(* IEC 61131-3 sources: sigmatek-logger-api/IXON_API/Network/IXON_Log, 1 file *)

(* ---- ONE_IXON_Log_Table.st ---- *)
#define OBJECTS_CONFIG

//Define part of class _TCPIPClient
#define TCPCLT_ERROR_NO            0
  #define TCPCLT_ERROR_INVALID_SOCK  -1
  #define TCPCLT_ERROR_CONNECTION    -2
  #define TCPCLT_ERROR_TIMEOUT       -3

  #define TCP_CLT_SEND_OK               0
  #define TCP_CLT_INVALID_HANDLE        -1
  #define TCP_CLT_NOT_CONNECTED         -2
  #define TCP_CLT_SEND_FAILED           -3
  #define TCP_CLT_SEND_BUFFER_FULL      -4
  #define TCP_CLT_DATA_TO_BIG_FOR_DIRECT_SENDING   -5
  #define TCP_CLT_MAXLEN_SEMANAME     32

  #define TCP_CLT_ERR_SET_PARA_INVALID_CMD     -10
  #define TCP_CLT_ERR_SET_PARA_INVALID_SUB_CMD -11

  #define TCP_CLT_ERR_TASK_ALREADY_EXIST       -12

  #define TCP_CLT_ERR_SET_PARA_CMD_NOT_SUPPORTED  -13

  #ifndef OS_VERSION_MIN_SALAMANDER
    #define OS_VERSION_MIN_SALAMANDER          0x9000
  #endif

  #define TCP_CLT_NO_ERROR                          0

  // - RETURN VALUES PRIVATE METHOD Read_LSLOBJ_CRC32
  #define TCP_CLT_ERR_GET_LSLOBJ_NAME             -20
  #define TCP_CLT_ERR_INVALID_POINTER             -21

  // - RETURN VALUES PRIVATE METHOD Read_AP_TaskPeriod
  #define TCP_CLT_ERR_TASK_TIME_NO_APP            -31
  #define TCP_CLT_ERR_TASK_TIME_WRONG_TASK_TYPE   -33
  #define TCP_CLT_ERR_TASK_TIME_OBJ_NOT_FOUND     -35

  // - RETURN VALUES PRIVATE METHOD AP_TaskCreate
  #define TCP_CLT_ERR_TASK_CREATE                 -40

  // - RETURN VALUES PRIVATE METHOD AP_SemaCreate
  #define TCP_CLT_ERR_SEMA_CREATE                 -50
  #define TCP_CLT_ERR_SEMA_INVALID_IDX            -51
  #define TCP_CLT_ERR_SEMA_INVALID_NAME           -52

  #define TCP_CLT_SEND_BUFFER_EMPTY                -6
  #define TCP_CLT_ERR_SEND_BUFFER_FATAL_ERROR      -7

  #define TCP_CLT_ERR_NO_SSL_INTERFACE             -8
  #define TCP_CLT_ERR_NO_TCP_INTERFACE             -9

  #define TCP_CLT_ERR_INVALID_PARA_TCP            -60
  #define TCP_CLT_ERR_INVALID_PARA_SSL            -61

  #define TCP_CLT_ERR_CONN_MEMORY                 -70
  #define TCP_CLT_ERR_MAX_CONN                    -80
  #define TCP_CLT_ERR_MAIN_INIT                   -90

  #define TCP_CLT_ERR_GROUP_OS                      0
  #define TCP_CLT_ERR_GROUP_AP                      1

  #define TCP_CLT_ERR_CODE_AP_TIMEOUT              -1

  #ifndef INIT_FIRSTSCAN
    #define INIT_FIRSTSCAN                         12
  #endif

  #ifndef AP_TASK_PRIORITY_DEFAULT
    #define AP_TASK_PRIORITY_DEFAULT               14
  #endif

  #define TCP_CLT_CMD_KEEP_ALIVE_PARA               2
  #define TCP_CLT_SUB_CMD_KEEP_ALIVE_INTERVAL       0
  #define TCP_CLT_SUB_CMD_KEEP_ALIVE_RETRY          1
  #define TCP_CLT_SUB_CMD_KEEP_ALIVE_TIMEOUT        2

  #define TCP_CLT_INFO_DISCONNECT                   0
  #define TCP_CLT_INFO_CONNECT                      1
  #define TCP_CLT_INFO_DELETED                      2

  #ifndef KEEPALIVE_INTERVAL_DEFAULT
    #define KEEPALIVE_INTERVAL_DEFAULT           7200
  #endif

  #ifndef KEEPALIVE_RETRYTIME_DEFAULT
    #define KEEPALIVE_RETRYTIME_DEFAULT            75
  #endif

  #ifndef KEEPALIVE_RETRYCNT_DEFUALT
    #define KEEPALIVE_RETRYCNT_DEFUALT             10
  #endif

  #ifndef CLOSE_SOCKET_TYPE_DEFAULT
    #define CLOSE_SOCKET_TYPE_DEFAULT               0
  #endif
#include "..\..\Class\_TCPIPClient\_TCPIPClient.h"
#include "..\..\Class\_TCPIPClient\SalamanderDelay.h"
#include "..\..\Class\_TCPIPClient\lsl_st_ssl_user.h"
//Define part of class cIXONConv10Value
#DEFINE MAX_NAME_LENGTH 100
#DEFINE MAX_VALUE_LENGTH 10
#DEFINE MAX_DATASTRING_LENGTH 1024
//Define part of class cIXONConv5Int5Str
#DEFINE MAX_NAME_LENGTH 100
#DEFINE MAX_INTEGER_LENGTH 10
#DEFINE MAX_DATASTRING_LENGTH 1024
#DEFINE MAX_STRING_LENGTH 100
//Define part of class IXON_LoggerAPI_Interface
#define SND_DATA_ARRAY_SIZE 1024
#define SND_ARRAY_SIZE 20
#define RCV_DATA_ARRAY_SIZE 1024
#include <.\lsl_st_mt.h>

FUNCTION GLOBAL TAB ONE_IXON_Log
-1$UINT, 0$UINT,
0$UINT, 0$UINT,

12$UDINT,
TO_UDINT(916194998), "_CheckSum", 1$UINT, 0$UINT, 1$UINT,
TO_UDINT(1778057824), "_TCPIPClient", 1$UINT, 1$UINT, 1$UINT,
TO_UDINT(670188634), "_TCPIPClientInterface", 1$UINT, 1$UINT, 0$UINT,
TO_UDINT(2199147857), "cIXONConv10Value", 0$UINT, 0$UINT, 1$UINT,
TO_UDINT(2966690256), "cIXONConv5Int5Str", 0$UINT, 0$UINT, 1$UINT,
TO_UDINT(2366984241), "IXON_LoggerAPI", 0$UINT, 0$UINT, 1$UINT,
TO_UDINT(357781282), "IXON_LoggerAPI_Interface", 0$UINT, 0$UINT, 1$UINT,
TO_UDINT(2225119864), "MerkerEx", 1$UINT, 22$UINT, 33$UINT,
TO_UDINT(3963750506), "Pulse", 0$UINT, 0$UINT, 1$UINT,
TO_UDINT(1850111279), "String", 1$UINT, 11$UINT, 33$UINT,
TO_UDINT(2898603620), "StringInternal", 1$UINT, 84$UINT, 0$UINT,
TO_UDINT(3232495061), "VirtualBaseInit", 1$UINT, 3$UINT, 0$UINT,

1$UINT, TO_UDINT(3180115317), "IXON_LOGGERAPI1\_TCPIPCLIENT1\CHECKSUM",

1$UINT, TO_UDINT(1796594274), "IXON_LOGGERAPI1\_TCPIPCLIENT1",

_NO_ATTR, TO_UDINT(3085999121), "GRIPPERSIXONLOG",

_NO_ATTR, TO_UDINT(1798062204), "BATCHIXONLOG",

_NO_ATTR, TO_UDINT(3532651229), "IXON_LOGGERAPI1",

1$UINT, TO_UDINT(1003265729), "IXON_LOGGERAPI1\MYTCPIPCLIENT1",

1$UINT, TO_UDINT(3192771373), "BATCHIXONLOG\INTEGERNAME1\MERKEREX0",
1$UINT, TO_UDINT(665826604), "BATCHIXONLOG\INTEGERNAME2\MERKEREX0",
1$UINT, TO_UDINT(3860949740), "BATCHIXONLOG\INTEGERNAME3\MERKEREX0",
1$UINT, TO_UDINT(3474620271), "BATCHIXONLOG\INTEGERNAME4\MERKEREX0",
1$UINT, TO_UDINT(244621487), "BATCHIXONLOG\INTEGERNAME5\MERKEREX0",
1$UINT, TO_UDINT(2181923968), "BATCHIXONLOG\STRING1\MERKEREX0",
1$UINT, TO_UDINT(468705921), "BATCHIXONLOG\STRING2\MERKEREX0",
1$UINT, TO_UDINT(3663805761), "BATCHIXONLOG\STRING3\MERKEREX0",
1$UINT, TO_UDINT(4082772162), "BATCHIXONLOG\STRING4\MERKEREX0",
1$UINT, TO_UDINT(852817666), "BATCHIXONLOG\STRING5\MERKEREX0",
1$UINT, TO_UDINT(2342531462), "BATCHIXONLOG\STRINGNAME1\MERKEREX0",
1$UINT, TO_UDINT(306337671), "BATCHIXONLOG\STRINGNAME2\MERKEREX0",
1$UINT, TO_UDINT(3553396807), "BATCHIXONLOG\STRINGNAME3\MERKEREX0",
1$UINT, TO_UDINT(4210531780), "BATCHIXONLOG\STRINGNAME4\MERKEREX0",
1$UINT, TO_UDINT(997802500), "BATCHIXONLOG\STRINGNAME5\MERKEREX0",
1$UINT, TO_UDINT(2779010355), "BATCHIXONLOG\TRIGGERNAME\MERKEREX0",
1$UINT, TO_UDINT(4245150780), "GRIPPERSIXONLOG\NAME10\MERKEREX0",
1$UINT, TO_UDINT(2566426530), "GRIPPERSIXONLOG\NAME1\MERKEREX0",
1$UINT, TO_UDINT(18540963), "GRIPPERSIXONLOG\NAME2\MERKEREX0",
1$UINT, TO_UDINT(3230938723), "GRIPPERSIXONLOG\NAME3\MERKEREX0",
1$UINT, TO_UDINT(3920569312), "GRIPPERSIXONLOG\NAME4\MERKEREX0",
1$UINT, TO_UDINT(673315872), "GRIPPERSIXONLOG\NAME5\MERKEREX0",
1$UINT, TO_UDINT(2982386209), "GRIPPERSIXONLOG\NAME6\MERKEREX0",
1$UINT, TO_UDINT(1884112353), "GRIPPERSIXONLOG\NAME7\MERKEREX0",
1$UINT, TO_UDINT(3820335399), "GRIPPERSIXONLOG\NAME8\MERKEREX0",
1$UINT, TO_UDINT(574320359), "GRIPPERSIXONLOG\NAME9\MERKEREX0",
1$UINT, TO_UDINT(3865678693), "GRIPPERSIXONLOG\TRIGGERNAME\MERKEREX0",
1$UINT, TO_UDINT(2981893656), "IXON_LOGGERAPI1\MYTCPIPCLIENT1\ST_IPADDRIXON\MERKEREX0",
1$UINT, TO_UDINT(2486479070), "IXON_LOGGERAPI1\MYTCPIPCLIENT1\ST_IPADDRPLC\MERKEREX0",
1$UINT, TO_UDINT(3086082301), "IXON_LOGGERAPI1\MYTCPIPCLIENT1\ST_PASSWORDIXON\MERKEREX0",
1$UINT, TO_UDINT(3369279868), "IXON_LOGGERAPI1\_TCPIPCLIENT1\STRSEMANAME01\MERKEREX0",
1$UINT, TO_UDINT(1362184061), "IXON_LOGGERAPI1\_TCPIPCLIENT1\STRSEMANAME02\MERKEREX0",
1$UINT, TO_UDINT(3451953391), "IXON_LOGGERAPI1\_TCPIPCLIENT1\STRTASKNAME\MERKEREX0",

_NO_ATTR, TO_UDINT(777463289), "PULSE1",

1$UINT, TO_UDINT(808633261), "BATCHIXONLOG\INTEGERNAME1",
1$UINT, TO_UDINT(2839253527), "BATCHIXONLOG\INTEGERNAME2",
1$UINT, TO_UDINT(3728515713), "BATCHIXONLOG\INTEGERNAME3",
1$UINT, TO_UDINT(1079523106), "BATCHIXONLOG\INTEGERNAME4",
1$UINT, TO_UDINT(928974772), "BATCHIXONLOG\INTEGERNAME5",
1$UINT, TO_UDINT(4091281586), "BATCHIXONLOG\STRING1",
1$UINT, TO_UDINT(1792364808), "BATCHIXONLOG\STRING2",
1$UINT, TO_UDINT(500326814), "BATCHIXONLOG\STRING3",
1$UINT, TO_UDINT(2209805373), "BATCHIXONLOG\STRING4",
1$UINT, TO_UDINT(4105290923), "BATCHIXONLOG\STRING5",
1$UINT, TO_UDINT(1673436439), "BATCHIXONLOG\STRINGNAME1",
1$UINT, TO_UDINT(4206349485), "BATCHIXONLOG\STRINGNAME2",
1$UINT, TO_UDINT(2377186363), "BATCHIXONLOG\STRINGNAME3",
1$UINT, TO_UDINT(332687768), "BATCHIXONLOG\STRINGNAME4",
1$UINT, TO_UDINT(1691572494), "BATCHIXONLOG\STRINGNAME5",
1$UINT, TO_UDINT(3473702409), "BATCHIXONLOG\TRIGGERNAME",
1$UINT, TO_UDINT(813494443), "GRIPPERSIXONLOG\NAME1",
1$UINT, TO_UDINT(3052394929), "GRIPPERSIXONLOG\NAME10",
1$UINT, TO_UDINT(2843058449), "GRIPPERSIXONLOG\NAME2",
1$UINT, TO_UDINT(3732050311), "GRIPPERSIXONLOG\NAME3",
1$UINT, TO_UDINT(1075184676), "GRIPPERSIXONLOG\NAME4",
1$UINT, TO_UDINT(923874482), "GRIPPERSIXONLOG\NAME5",
1$UINT, TO_UDINT(2920834312), "GRIPPERSIXONLOG\NAME6",
1$UINT, TO_UDINT(3642709406), "GRIPPERSIXONLOG\NAME7",
1$UINT, TO_UDINT(1235240975), "GRIPPERSIXONLOG\NAME8",
1$UINT, TO_UDINT(1051162777), "GRIPPERSIXONLOG\NAME9",
1$UINT, TO_UDINT(3416962169), "GRIPPERSIXONLOG\TRIGGERNAME",
1$UINT, TO_UDINT(2721538750), "IXON_LOGGERAPI1\MYTCPIPCLIENT1\ST_IPADDRIXON",
1$UINT, TO_UDINT(1805041610), "IXON_LOGGERAPI1\MYTCPIPCLIENT1\ST_IPADDRPLC",
1$UINT, TO_UDINT(1852407263), "IXON_LOGGERAPI1\MYTCPIPCLIENT1\ST_PASSWORDIXON",
1$UINT, TO_UDINT(962394143), "IXON_LOGGERAPI1\_TCPIPCLIENT1\STRSEMANAME01",
1$UINT, TO_UDINT(2689968549), "IXON_LOGGERAPI1\_TCPIPCLIENT1\STRSEMANAME02",
1$UINT, TO_UDINT(2790321702), "IXON_LOGGERAPI1\_TCPIPCLIENT1\STRTASKNAME",

//Internal connections
0$UDINT,
69$UDINT,
TO_UDINT(1), "CheckSum", TO_UDINT(0),
TO_UDINT(1), "StrTaskName", TO_UDINT(72),
TO_UDINT(1), "StrSemaName01", TO_UDINT(70),
TO_UDINT(1), "StrSemaName02", TO_UDINT(71),
TO_UDINT(2), "Name3", TO_UDINT(59),
TO_UDINT(2), "Name2", TO_UDINT(58),
TO_UDINT(2), "Name1", TO_UDINT(56),
TO_UDINT(2), "Name4", TO_UDINT(60),
TO_UDINT(2), "Name5", TO_UDINT(61),
TO_UDINT(2), "Name6", TO_UDINT(62),
TO_UDINT(2), "Name7", TO_UDINT(63),
TO_UDINT(2), "Name8", TO_UDINT(64),
TO_UDINT(2), "Name9", TO_UDINT(65),
TO_UDINT(2), "Name10", TO_UDINT(57),
TO_UDINT(2), "TriggerName", TO_UDINT(66),
TO_UDINT(3), "TriggerName", TO_UDINT(55),
TO_UDINT(3), "String1", TO_UDINT(45),
TO_UDINT(3), "String2", TO_UDINT(46),
TO_UDINT(3), "String3", TO_UDINT(47),
TO_UDINT(3), "String4", TO_UDINT(48),
TO_UDINT(3), "String5", TO_UDINT(49),
TO_UDINT(3), "IntegerName1", TO_UDINT(40),
TO_UDINT(3), "IntegerName2", TO_UDINT(41),
TO_UDINT(3), "IntegerName3", TO_UDINT(42),
TO_UDINT(3), "IntegerName4", TO_UDINT(43),
TO_UDINT(3), "IntegerName5", TO_UDINT(44),
TO_UDINT(3), "StringName1", TO_UDINT(50),
TO_UDINT(3), "StringName2", TO_UDINT(51),
TO_UDINT(3), "StringName3", TO_UDINT(52),
TO_UDINT(3), "StringName4", TO_UDINT(53),
TO_UDINT(3), "StringName5", TO_UDINT(54),
TO_UDINT(4), "_TCPIPClient1", TO_UDINT(1),
TO_UDINT(4), "MyTCPIPClient1", TO_UDINT(5),
TO_UDINT(5), "ST_IPAddrIXON", TO_UDINT(67),
TO_UDINT(5), "ST_PasswordIXON", TO_UDINT(69),
TO_UDINT(5), "ST_IPAddrPLC", TO_UDINT(68),
TO_UDINT(40), "MerkerEx0", TO_UDINT(6),
TO_UDINT(41), "MerkerEx0", TO_UDINT(7),
TO_UDINT(42), "MerkerEx0", TO_UDINT(8),
TO_UDINT(43), "MerkerEx0", TO_UDINT(9),
TO_UDINT(44), "MerkerEx0", TO_UDINT(10),
TO_UDINT(45), "MerkerEx0", TO_UDINT(11),
TO_UDINT(46), "MerkerEx0", TO_UDINT(12),
TO_UDINT(47), "MerkerEx0", TO_UDINT(13),
TO_UDINT(48), "MerkerEx0", TO_UDINT(14),
TO_UDINT(49), "MerkerEx0", TO_UDINT(15),
TO_UDINT(50), "MerkerEx0", TO_UDINT(16),
TO_UDINT(51), "MerkerEx0", TO_UDINT(17),
TO_UDINT(52), "MerkerEx0", TO_UDINT(18),
TO_UDINT(53), "MerkerEx0", TO_UDINT(19),
TO_UDINT(54), "MerkerEx0", TO_UDINT(20),
TO_UDINT(55), "MerkerEx0", TO_UDINT(21),
TO_UDINT(56), "MerkerEx0", TO_UDINT(23),
TO_UDINT(57), "MerkerEx0", TO_UDINT(22),
TO_UDINT(58), "MerkerEx0", TO_UDINT(24),
TO_UDINT(59), "MerkerEx0", TO_UDINT(25),
TO_UDINT(60), "MerkerEx0", TO_UDINT(26),
TO_UDINT(61), "MerkerEx0", TO_UDINT(27),
TO_UDINT(62), "MerkerEx0", TO_UDINT(28),
TO_UDINT(63), "MerkerEx0", TO_UDINT(29),
TO_UDINT(64), "MerkerEx0", TO_UDINT(30),
TO_UDINT(65), "MerkerEx0", TO_UDINT(31),
TO_UDINT(66), "MerkerEx0", TO_UDINT(32),
TO_UDINT(67), "MerkerEx0", TO_UDINT(33),
TO_UDINT(68), "MerkerEx0", TO_UDINT(34),
TO_UDINT(69), "MerkerEx0", TO_UDINT(35),
TO_UDINT(70), "MerkerEx0", TO_UDINT(36),
TO_UDINT(71), "MerkerEx0", TO_UDINT(37),
TO_UDINT(72), "MerkerEx0", TO_UDINT(38),
0$UDINT,
39$UDINT,
TO_UDINT(2), "ToIXON_LoggerAPI", TO_UDINT(5), "ClassSvr",
TO_UDINT(3), "ToIXON_LoggerAPI", TO_UDINT(5), "ClassSvr",
TO_UDINT(5), "_TCPIPClient", TO_UDINT(1), "Control",
TO_UDINT(39), "PulseOut1", TO_UDINT(2), "sCmdConvert",
TO_UDINT(39), "PulseOut2", TO_UDINT(2), "sValue1",
TO_UDINT(39), "PulseOut3", TO_UDINT(3), "sCmdConvert",
TO_UDINT(40), "DataBuffer", TO_UDINT(6), "m_udLength",
TO_UDINT(41), "DataBuffer", TO_UDINT(7), "m_udLength",
TO_UDINT(42), "DataBuffer", TO_UDINT(8), "m_udLength",
TO_UDINT(43), "DataBuffer", TO_UDINT(9), "m_udLength",
TO_UDINT(44), "DataBuffer", TO_UDINT(10), "m_udLength",
TO_UDINT(45), "DataBuffer", TO_UDINT(11), "m_udLength",
TO_UDINT(46), "DataBuffer", TO_UDINT(12), "m_udLength",
TO_UDINT(47), "DataBuffer", TO_UDINT(13), "m_udLength",
TO_UDINT(48), "DataBuffer", TO_UDINT(14), "m_udLength",
TO_UDINT(49), "DataBuffer", TO_UDINT(15), "m_udLength",
TO_UDINT(50), "DataBuffer", TO_UDINT(16), "m_udLength",
TO_UDINT(51), "DataBuffer", TO_UDINT(17), "m_udLength",
TO_UDINT(52), "DataBuffer", TO_UDINT(18), "m_udLength",
TO_UDINT(53), "DataBuffer", TO_UDINT(19), "m_udLength",
TO_UDINT(54), "DataBuffer", TO_UDINT(20), "m_udLength",
TO_UDINT(55), "DataBuffer", TO_UDINT(21), "m_udLength",
TO_UDINT(56), "DataBuffer", TO_UDINT(23), "m_udLength",
TO_UDINT(57), "DataBuffer", TO_UDINT(22), "m_udLength",
TO_UDINT(58), "DataBuffer", TO_UDINT(24), "m_udLength",
TO_UDINT(59), "DataBuffer", TO_UDINT(25), "m_udLength",
TO_UDINT(60), "DataBuffer", TO_UDINT(26), "m_udLength",
TO_UDINT(61), "DataBuffer", TO_UDINT(27), "m_udLength",
TO_UDINT(62), "DataBuffer", TO_UDINT(28), "m_udLength",
TO_UDINT(63), "DataBuffer", TO_UDINT(29), "m_udLength",
TO_UDINT(64), "DataBuffer", TO_UDINT(30), "m_udLength",
TO_UDINT(65), "DataBuffer", TO_UDINT(31), "m_udLength",
TO_UDINT(66), "DataBuffer", TO_UDINT(32), "m_udLength",
TO_UDINT(67), "DataBuffer", TO_UDINT(33), "m_udLength",
TO_UDINT(68), "DataBuffer", TO_UDINT(34), "m_udLength",
TO_UDINT(69), "DataBuffer", TO_UDINT(35), "m_udLength",
TO_UDINT(70), "DataBuffer", TO_UDINT(36), "m_udLength",
TO_UDINT(71), "DataBuffer", TO_UDINT(37), "m_udLength",
TO_UDINT(72), "DataBuffer", TO_UDINT(38), "m_udLength",

//Initialization values
0$UDINT,
71$UDINT,
TO_UDINT(1), "Port", TO_UDINT(9230),//|IXON_Log.IXON_LoggerAPI1\_TCPIPClient1.Port;
TO_UDINT(1), "MaxConnections", TO_UDINT(0),//|IXON_Log.IXON_LoggerAPI1\_TCPIPClient1.MaxConnections;
TO_UDINT(2), "sSetInitNrOfEntrys", TO_UDINT(8),//|IXON_Log.GrippersIXONLog.sSetInitNrOfEntrys;
TO_UDINT(3), "sSetInitNrOfInteger", TO_UDINT(1),//|IXON_Log.BatchIXONLog.sSetInitNrOfInteger;
TO_UDINT(3), "sSetInitNrOfString", TO_UDINT(3),//|IXON_Log.BatchIXONLog.sSetInitNrOfString;
TO_UDINT(6), "ThreadSafe", TO_UDINT(0),//|IXON_Log.IntegerName1\BatchIXONLog\MerkerEx0.ThreadSafe;
TO_UDINT(7), "ThreadSafe", TO_UDINT(0),//|IXON_Log.IntegerName2\BatchIXONLog\MerkerEx0.ThreadSafe;
TO_UDINT(8), "ThreadSafe", TO_UDINT(0),//|IXON_Log.IntegerName3\BatchIXONLog\MerkerEx0.ThreadSafe;
TO_UDINT(9), "ThreadSafe", TO_UDINT(0),//|IXON_Log.IntegerName4\BatchIXONLog\MerkerEx0.ThreadSafe;
TO_UDINT(10), "ThreadSafe", TO_UDINT(0),//|IXON_Log.IntegerName5\BatchIXONLog\MerkerEx0.ThreadSafe;
TO_UDINT(11), "ThreadSafe", TO_UDINT(0),//|IXON_Log.String1\BatchIXONLog\MerkerEx0.ThreadSafe;
TO_UDINT(12), "ThreadSafe", TO_UDINT(0),//|IXON_Log.String2\BatchIXONLog\MerkerEx0.ThreadSafe;
TO_UDINT(13), "ThreadSafe", TO_UDINT(0),//|IXON_Log.String3\BatchIXONLog\MerkerEx0.ThreadSafe;
TO_UDINT(14), "ThreadSafe", TO_UDINT(0),//|IXON_Log.String4\BatchIXONLog\MerkerEx0.ThreadSafe;
TO_UDINT(15), "ThreadSafe", TO_UDINT(0),//|IXON_Log.String5\BatchIXONLog\MerkerEx0.ThreadSafe;
TO_UDINT(16), "ThreadSafe", TO_UDINT(0),//|IXON_Log.StringName1\BatchIXONLog\MerkerEx0.ThreadSafe;
TO_UDINT(17), "ThreadSafe", TO_UDINT(0),//|IXON_Log.StringName2\BatchIXONLog\MerkerEx0.ThreadSafe;
TO_UDINT(18), "ThreadSafe", TO_UDINT(0),//|IXON_Log.StringName3\BatchIXONLog\MerkerEx0.ThreadSafe;
TO_UDINT(19), "ThreadSafe", TO_UDINT(0),//|IXON_Log.StringName4\BatchIXONLog\MerkerEx0.ThreadSafe;
TO_UDINT(20), "ThreadSafe", TO_UDINT(0),//|IXON_Log.StringName5\BatchIXONLog\MerkerEx0.ThreadSafe;
TO_UDINT(21), "ThreadSafe", TO_UDINT(0),//|IXON_Log.TriggerName\BatchIXONLog\MerkerEx0.ThreadSafe;
TO_UDINT(22), "ThreadSafe", TO_UDINT(0),//|IXON_Log.Name10\GrippersIXONLog\MerkerEx0.ThreadSafe;
TO_UDINT(23), "ThreadSafe", TO_UDINT(0),//|IXON_Log.Name1\GrippersIXONLog\MerkerEx0.ThreadSafe;
TO_UDINT(24), "ThreadSafe", TO_UDINT(0),//|IXON_Log.Name2\GrippersIXONLog\MerkerEx0.ThreadSafe;
TO_UDINT(25), "ThreadSafe", TO_UDINT(0),//|IXON_Log.Name3\GrippersIXONLog\MerkerEx0.ThreadSafe;
TO_UDINT(26), "ThreadSafe", TO_UDINT(0),//|IXON_Log.Name4\GrippersIXONLog\MerkerEx0.ThreadSafe;
TO_UDINT(27), "ThreadSafe", TO_UDINT(0),//|IXON_Log.Name5\GrippersIXONLog\MerkerEx0.ThreadSafe;
TO_UDINT(28), "ThreadSafe", TO_UDINT(0),//|IXON_Log.Name6\GrippersIXONLog\MerkerEx0.ThreadSafe;
TO_UDINT(29), "ThreadSafe", TO_UDINT(0),//|IXON_Log.Name7\GrippersIXONLog\MerkerEx0.ThreadSafe;
TO_UDINT(30), "ThreadSafe", TO_UDINT(0),//|IXON_Log.Name8\GrippersIXONLog\MerkerEx0.ThreadSafe;
TO_UDINT(31), "ThreadSafe", TO_UDINT(0),//|IXON_Log.Name9\GrippersIXONLog\MerkerEx0.ThreadSafe;
TO_UDINT(32), "ThreadSafe", TO_UDINT(0),//|IXON_Log.TriggerName\GrippersIXONLog\MerkerEx0.ThreadSafe;
TO_UDINT(33), "ThreadSafe", TO_UDINT(0),//|IXON_Log.ST_IPAddrIXON\MyTCPIPClient1\IXON_LoggerAPI1\MerkerEx0.ThreadSafe;
TO_UDINT(34), "ThreadSafe", TO_UDINT(0),//|IXON_Log.ST_IPAddrPLC\MyTCPIPClient1\IXON_LoggerAPI1\MerkerEx0.ThreadSafe;
TO_UDINT(35), "ThreadSafe", TO_UDINT(0),//|IXON_Log.ST_PasswordIXON\MyTCPIPClient1\IXON_LoggerAPI1\MerkerEx0.ThreadSafe;
TO_UDINT(36), "ThreadSafe", TO_UDINT(0),//|IXON_Log.StrSemaName01\_TCPIPClient1\IXON_LoggerAPI1\MerkerEx0.ThreadSafe;
TO_UDINT(37), "ThreadSafe", TO_UDINT(0),//|IXON_Log.StrSemaName02\_TCPIPClient1\IXON_LoggerAPI1\MerkerEx0.ThreadSafe;
TO_UDINT(38), "ThreadSafe", TO_UDINT(0),//|IXON_Log.StrTaskName\_TCPIPClient1\IXON_LoggerAPI1\MerkerEx0.ThreadSafe;
TO_UDINT(40), "SingleRealloc", TO_UDINT(1),//|IXON_Log.BatchIXONLog\IntegerName1.SingleRealloc;
TO_UDINT(41), "SingleRealloc", TO_UDINT(1),//|IXON_Log.BatchIXONLog\IntegerName2.SingleRealloc;
TO_UDINT(42), "SingleRealloc", TO_UDINT(1),//|IXON_Log.BatchIXONLog\IntegerName3.SingleRealloc;
TO_UDINT(43), "SingleRealloc", TO_UDINT(1),//|IXON_Log.BatchIXONLog\IntegerName4.SingleRealloc;
TO_UDINT(44), "SingleRealloc", TO_UDINT(1),//|IXON_Log.BatchIXONLog\IntegerName5.SingleRealloc;
TO_UDINT(45), "SingleRealloc", TO_UDINT(1),//|IXON_Log.BatchIXONLog\String1.SingleRealloc;
TO_UDINT(46), "SingleRealloc", TO_UDINT(1),//|IXON_Log.BatchIXONLog\String2.SingleRealloc;
TO_UDINT(47), "SingleRealloc", TO_UDINT(1),//|IXON_Log.BatchIXONLog\String3.SingleRealloc;
TO_UDINT(48), "SingleRealloc", TO_UDINT(1),//|IXON_Log.BatchIXONLog\String4.SingleRealloc;
TO_UDINT(49), "SingleRealloc", TO_UDINT(1),//|IXON_Log.BatchIXONLog\String5.SingleRealloc;
TO_UDINT(50), "SingleRealloc", TO_UDINT(1),//|IXON_Log.BatchIXONLog\StringName1.SingleRealloc;
TO_UDINT(51), "SingleRealloc", TO_UDINT(1),//|IXON_Log.BatchIXONLog\StringName2.SingleRealloc;
TO_UDINT(52), "SingleRealloc", TO_UDINT(1),//|IXON_Log.BatchIXONLog\StringName3.SingleRealloc;
TO_UDINT(53), "SingleRealloc", TO_UDINT(1),//|IXON_Log.BatchIXONLog\StringName4.SingleRealloc;
TO_UDINT(54), "SingleRealloc", TO_UDINT(1),//|IXON_Log.BatchIXONLog\StringName5.SingleRealloc;
TO_UDINT(55), "SingleRealloc", TO_UDINT(1),//|IXON_Log.BatchIXONLog\TriggerName.SingleRealloc;
TO_UDINT(56), "SingleRealloc", TO_UDINT(1),//|IXON_Log.GrippersIXONLog\Name1.SingleRealloc;
TO_UDINT(57), "SingleRealloc", TO_UDINT(1),//|IXON_Log.GrippersIXONLog\Name10.SingleRealloc;
TO_UDINT(58), "SingleRealloc", TO_UDINT(1),//|IXON_Log.GrippersIXONLog\Name2.SingleRealloc;
TO_UDINT(59), "SingleRealloc", TO_UDINT(1),//|IXON_Log.GrippersIXONLog\Name3.SingleRealloc;
TO_UDINT(60), "SingleRealloc", TO_UDINT(1),//|IXON_Log.GrippersIXONLog\Name4.SingleRealloc;
TO_UDINT(61), "SingleRealloc", TO_UDINT(1),//|IXON_Log.GrippersIXONLog\Name5.SingleRealloc;
TO_UDINT(62), "SingleRealloc", TO_UDINT(1),//|IXON_Log.GrippersIXONLog\Name6.SingleRealloc;
TO_UDINT(63), "SingleRealloc", TO_UDINT(1),//|IXON_Log.GrippersIXONLog\Name7.SingleRealloc;
TO_UDINT(64), "SingleRealloc", TO_UDINT(1),//|IXON_Log.GrippersIXONLog\Name8.SingleRealloc;
TO_UDINT(65), "SingleRealloc", TO_UDINT(1),//|IXON_Log.GrippersIXONLog\Name9.SingleRealloc;
TO_UDINT(66), "SingleRealloc", TO_UDINT(1),//|IXON_Log.GrippersIXONLog\TriggerName.SingleRealloc;
TO_UDINT(67), "SingleRealloc", TO_UDINT(1),//|IXON_Log.MyTCPIPClient1\IXON_LoggerAPI1\ST_IPAddrIXON.SingleRealloc;
TO_UDINT(68), "SingleRealloc", TO_UDINT(1),//|IXON_Log.MyTCPIPClient1\IXON_LoggerAPI1\ST_IPAddrPLC.SingleRealloc;
TO_UDINT(69), "SingleRealloc", TO_UDINT(1),//|IXON_Log.MyTCPIPClient1\IXON_LoggerAPI1\ST_PasswordIXON.SingleRealloc;
TO_UDINT(70), "SingleRealloc", TO_UDINT(1),//|IXON_Log._TCPIPClient1\IXON_LoggerAPI1\StrSemaName01.SingleRealloc;
TO_UDINT(71), "SingleRealloc", TO_UDINT(1),//|IXON_Log._TCPIPClient1\IXON_LoggerAPI1\StrSemaName02.SingleRealloc;
TO_UDINT(72), "SingleRealloc", TO_UDINT(1),//|IXON_Log._TCPIPClient1\IXON_LoggerAPI1\StrTaskName.SingleRealloc;

//Symbolic initialization values
0$UDINT,
0$UDINT,

//Initialization of string values
0$UDINT,
22$UDINT,
TO_UDINT(40), "", 0$UINT, TO_UINT(OFF(L1)-OFF(L0)), L0:"NrOfPlantingCycles",L1://|IXON_Log.BatchIXONLog\IntegerName1.Data;
TO_UDINT(45), "", 0$UINT, TO_UINT(OFF(L3)-OFF(L2)), L2:"2022-01-07 10:45:21",L3://|IXON_Log.BatchIXONLog\String1.Data;
TO_UDINT(46), "", 0$UINT, TO_UINT(OFF(L5)-OFF(L4)), L4:"2022-01-07 11:09:21",L5://|IXON_Log.BatchIXONLog\String2.Data;
TO_UDINT(47), "", 0$UINT, TO_UINT(OFF(L7)-OFF(L6)), L6:"Batch 123",L7://|IXON_Log.BatchIXONLog\String3.Data;
TO_UDINT(48), "", 0$UINT, TO_UINT(OFF(L9)-OFF(L8)), L8:1,L9://|IXON_Log.BatchIXONLog\String4.Data;
TO_UDINT(49), "", 0$UINT, TO_UINT(OFF(L11)-OFF(L10)), L10:0,L11://|IXON_Log.BatchIXONLog\String5.Data;
TO_UDINT(50), "", 0$UINT, TO_UINT(OFF(L13)-OFF(L12)), L12:"StartBatch",L13://|IXON_Log.BatchIXONLog\StringName1.Data;
TO_UDINT(51), "", 0$UINT, TO_UINT(OFF(L15)-OFF(L14)), L14:"EndBatch",L15://|IXON_Log.BatchIXONLog\StringName2.Data;
TO_UDINT(52), "", 0$UINT, TO_UINT(OFF(L17)-OFF(L16)), L16:"BatchName",L17://|IXON_Log.BatchIXONLog\StringName3.Data;
TO_UDINT(55), "", 0$UINT, TO_UINT(OFF(L19)-OFF(L18)), L18:"TrigBatch",L19://|IXON_Log.BatchIXONLog\TriggerName.Data;
TO_UDINT(56), "", 0$UINT, TO_UINT(OFF(L21)-OFF(L20)), L20:"LastGripperWithCommError",L21://|IXON_Log.GrippersIXONLog\Name1.Data;
TO_UDINT(58), "", 0$UINT, TO_UINT(OFF(L23)-OFF(L22)), L22:"NrOfCommErrors",L23://|IXON_Log.GrippersIXONLog\Name2.Data;
TO_UDINT(59), "", 0$UINT, TO_UINT(OFF(L25)-OFF(L24)), L24:0"GDSError",L25://|IXON_Log.GrippersIXONLog\Name3.Data;
TO_UDINT(60), "", 0$UINT, TO_UINT(OFF(L27)-OFF(L26)), L26:"OFFError",L27://|IXON_Log.GrippersIXONLog\Name4.Data;
TO_UDINT(61), "", 0$UINT, TO_UINT(OFF(L29)-OFF(L28)), L28:"MoveRetries",L29://|IXON_Log.GrippersIXONLog\Name5.Data;
TO_UDINT(62), "", 0$UINT, TO_UINT(OFF(L31)-OFF(L30)), L30:"NrOfTeaching",L31://|IXON_Log.GrippersIXONLog\Name6.Data;
TO_UDINT(63), "", 0$UINT, TO_UINT(OFF(L33)-OFF(L32)), L32:"GripperWithBiggestPosDiff",L33://|IXON_Log.GrippersIXONLog\Name7.Data;
TO_UDINT(64), "", 0$UINT, TO_UINT(OFF(L35)-OFF(L34)), L34:"TeachingPosDifference",L35://|IXON_Log.GrippersIXONLog\Name8.Data;
TO_UDINT(66), "", 0$UINT, TO_UINT(OFF(L37)-OFF(L36)), L36:"TrigGrippers",L37://|IXON_Log.GrippersIXONLog\TriggerName.Data;
TO_UDINT(67), "", 0$UINT, TO_UINT(OFF(L39)-OFF(L38)), L38:"192.168.150.1",L39://|IXON_Log.MyTCPIPClient1\IXON_LoggerAPI1\ST_IPAddrIXON.Data;
TO_UDINT(68), "", 0$UINT, TO_UINT(OFF(L41)-OFF(L40)), L40:"192.168.150.10",L41://|IXON_Log.MyTCPIPClient1\IXON_LoggerAPI1\ST_IPAddrPLC.Data;
TO_UDINT(69), "", 0$UINT, TO_UINT(OFF(L43)-OFF(L42)), L42:"1234",L43://|IXON_Log.MyTCPIPClient1\IXON_LoggerAPI1\ST_PasswordIXON.Data;

//Configuration of tasks (RealTime, Cyclic, Background)
0$UDINT,
0$UDINT,

0$UDINT,
3$UDINT,
TO_UDINT(1), (10)$UDINT, 4194303$DINT, 	//IXON_LOGGERAPI1\_TCPIPCLIENT1
TO_UDINT(5), (10)$UDINT, 4194303$DINT, 	//IXON_LOGGERAPI1\MYTCPIPCLIENT1
TO_UDINT(39), (500)$UDINT, 4194303$DINT, 	//PULSE1

0$UDINT,
0$UDINT,

//External connections
0$UDINT,
0$UDINT,

//Magic internal connections
0$UDINT,
0$UDINT,

//Configuration of timeslots of tasks (RealTime, Cyclic)
#ifdef __LSLLDR_TIMESLOTS__
0$UDINT,
0$UDINT,

0$UDINT,
0$UDINT,

#endif //__LSLLDR_TIMESLOTS__

//MultiMaster connections
#ifdef __LSLLDR_MULTIMASTER__
0$UDINT,
0$UDINT,
#endif //__LSLLDR_MULTIMASTER__

//Configuration for task ID (RealTime, CyclicTime)
#ifdef __LSLLDR_TASKID__
"\\\\TASKS2  "
0$UDINT,
0$UDINT,

0$UDINT,
3$UDINT,
(0)$UDINT, 	//IXON_LOGGERAPI1\_TCPIPCLIENT1
(0)$UDINT, 	//IXON_LOGGERAPI1\MYTCPIPCLIENT1
(0)$UDINT, 	//PULSE1

0$UDINT,
0$UDINT,

#endif //__LSLLDR_TASKID__

END_FUNCTION
